Yaskawa INFORM job: 1.JBI

/JOB
//NAME 1
//POS
///NPOS 162,162,162,0,0,0
///TOOL 0
///POSTYPE PULSE
///PULSE
C00000=-283,-101162,-84213,3710,-80188,-1936
C00001=-283,-101162,-84213,3710,-80188,-1936
C00002=115939,-17843,-44700,-6904,-63515,59085
C00003=117709,3731,-51645,-6384,-54030,83191
C00004=117709,3731,-51645,-6384,-54030,83191
C00005=124817,11091,-45240,2225,-58232,65802
C00006=128558,-4341,-61499,8943,-39416,48451
C00007=141937,23059,-44881,39121,-57053,20454
C00008=142920,35333,-35255,42486,-63609,8178
C00009=131389,51659,-10555,16038,-74664,11710
C00010=126196,50041,-9511,12612,-72523,-6101
C00011=114039,49083,-11086,-6822,-73270,-17046
C00012=112111,54426,-8133,-7185,-80829,-32375
C00013=101553,48559,-20697,-28143,-77568,-33966
C00014=105123,31884,-31701,-21046,-69946,-46894
C00015=111650,18447,-39836,-11003,-63489,-61522
C00016=113485,7970,-48571,-14105,-57851,-74639
C00017=113485,7970,-48571,-14105,-57851,-74639
C00018=114170,-2374,-36949,-11645,-74681,-76938
C00019=113314,-7643,-38017,-11019,-76954,88145
C00020=102960,15783,-40712,-5055,-61801,87407
C00021=102960,15783,-40712,-5055,-61801,87407
C00022=109484,11848,-44448,3017,-57913,70801
C00023=111825,-4491,-61766,4155,-38221,55572
C00024=127233,18004,-49993,42137,-51406,23800
C00025=123794,20070,-44223,34245,-49783,15146
C00026=118261,52920,-9530,17828,-74428,15725
C00027=113721,45593,-13485,15354,-67043,-2855
C00028=99817,50806,-8879,-9234,-71758,-11440
C00029=100311,60695,-910,-3132,-82683,-29064
C00030=89808,58501,-9489,-23508,-82083,-31436
C00031=93781,55410,-9430,-14151,-84882,-46382
C00032=94766,20128,-39423,-16116,-61452,-54210
C00033=98573,11657,-45494,-13692,-58332,-69623
C00034=98573,11657,-45494,-13692,-58332,-69623
C00035=99303,8604,-31154,-10952,-72489,-71699
C00036=89422,16015,-23794,-2157,-75183,91094
C00037=90041,28841,-28187,-2386,-65884,91066
C00038=90041,28841,-28187,-2386,-65884,91066
C00039=95426,19332,-37606,3682,-57792,75417
C00040=103247,16005,-44070,17550,-50613,56089
C00041=113549,16841,-53361,50996,-44891,24333
C00042=112114,26764,-40359,41262,-49930,18196
C00043=105423,50717,-10337,19910,-67719,16523
C00044=102098,58112,-1142,17447,-71662,1302
C00045=90776,64198,5929,-1117,-76945,-10230
C00046=87727,74947,14485,-3611,-87418,-24219
C00047=79354,72723,7405,-19240,-87200,-29236
C00048=76420,55305,-10510,-24564,-76474,-35505
C00049=83670,16895,-41951,-12582,-49930,-51607
C00050=85054,23740,-34298,-12468,-60756,-65460
C00051=85054,23740,-34298,-12468,-60756,-65460
C00052=85063,22114,-18753,-9149,-74798,-67250
C00053=72786,31521,-9549,-9445,-75352,93043
C00054=77617,39381,-17527,-2945,-63917,95499
C00055=77617,39381,-17527,-2945,-63917,95499
C00056=81845,27264,-30649,1079,-52677,78149
C00057=86990,13258,-48946,12655,-33027,60150
C00058=90994,9633,-56784,33436,-24362,42962
C00059=99247,25142,-45272,51284,-40942,28841
C00060=98491,33379,-33635,41928,-45438,21477
C00061=97892,43719,-21091,40448,-51711,6672
C00062=90154,66189,8945,17735,-69591,4970
C00063=76670,80759,24898,-8994,-81212,-4057
C00064=77890,93073,36819,-863,-92684,-21133
C00065=70280,91760,31185,-15532,-93504,-27367
C00066=65704,69069,5703,-24854,-77527,-31557
C00067=69263,47501,-12611,-17938,-65429,-45438
C00068=73833,39987,-17909,-11044,-63928,-62173
C00069=73833,39987,-17909,-11044,-63928,-62173
C00070=75039,37514,-3449,-7701,-77257,-64173
C00071=74616,28156,-12897,-9694,-74827,92488
C00072=73614,40170,-17462,-11390,-64426,94165
C00073=73614,40170,-17462,-11390,-64426,94165
C00074=73614,40170,-17462,-11390,-64426,94165
C00075=81727,26723,-31141,1076,-52650,80628
C00076=86883,12521,-49454,12588,-33076,60218
C00077=90994,9713,-56809,33527,-24311,42932
C00078=90994,9713,-56809,33527,-24311,42932
C00079=99183,24902,-45504,51304,-40911,28852
C00080=99183,24902,-45504,51304,-40911,28852
C00081=98411,33440,-33412,41862,-45487,21541
C00082=99416,42526,-24620,46864,-51095,3725
C00083=90863,70401,13127,18633,-73267,4997
C00084=76675,81176,25590,-8988,-81419,-4073
C00085=77890,93045,36838,-863,-92708,-21133
C00086=70280,91719,31202,-15533,-93535,-27371
C00087=65715,68855,5477,-24835,-77499,-31559
C00088=66119,47846,-14846,-25675,-64947,-43795
C00089=70910,45228,-13849,-14534,-65052,-50806
C00090=75926,27198,-30687,-6609,-51803,-64018
C00091=75926,27198,-30687,-6609,-51803,-64018
C00092=74844,35432,-1015,-7610,-79822,-64270
C00093=74616,28156,-12897,-9694,-74827,92488
C00094=90411,-2677,-20047,-11125,-84138,86440
C00095=90413,-2674,-20051,-11105,-84138,86441
C00096=137757,-12075,-30464,2646,-72394,74401
C00097=139263,-65150,-85436,14259,-28990,73053
C00098=137079,-26031,-69593,36686,-11816,62677
C00099=137079,-26031,-69593,36686,-11816,62677
C00100=139435,-23870,-66142,38084,-15914,40453
C00101=138383,-26116,-69231,45202,-10210,18865
C00102=136988,-21816,-61713,19512,-16285,9124
C00103=134481,-8714,-45390,4049,-32022,-3278
C00104=132816,-12054,-49266,2863,-29473,-26222
C00105=133118,-16915,-54850,5104,-25691,-47193
C00106=132429,-23928,-65383,-2979,-14980,-66671
C00107=133899,-27903,-74314,23479,-2636,-94546
C00108=138833,-79965,-103111,19688,-12213,-93629
C00109=119564,-93872,-103655,-3232,-19191,84847
C00110=119617,-28274,-68464,-3848,-15128,84753
C00111=119617,-28274,-68464,-3848,-15128,84753
C00112=119575,-30245,-73045,-30117,-7907,72568
C00113=119533,-30199,-72935,-30139,-8105,72141
C00114=119084,-28019,-67713,-21117,-14338,49832
C00115=119103,-25674,-64433,-15990,-16239,28421
C00116=117904,-24651,-63335,-18016,-16610,10465
C00117=116364,-17323,-54707,-12430,-26691,-16379
C00118=116034,-19270,-56740,-12888,-26506,-35915
C00119=108922,-18911,-60992,-47912,-30029,-42936
C00120=114993,-30399,-76205,-74620,-10810,-47413
C00121=113126,-78683,-102705,-45607,-16425,-60367
C00122=119564,-93872,-103655,-3232,-19191,84847
C00123=119501,-30079,-72867,-7033,-8758,86614
C00124=119501,-30079,-72867,-7033,-8758,86614
C00125=119390,-30716,-74067,-37591,-7172,75727
C00126=121229,-29061,-69555,-4595,-11344,43979
C00127=119104,-25703,-64453,-15989,-16243,28419
C00128=118126,-13614,-49952,-9217,-30446,5536
C00129=116206,-13809,-50361,-10582,-31136,-17197
C00130=117334,-18567,-55575,-6506,-27346,-35991
C00131=112042,-24638,-66931,-46893,-21308,-43852
C00132=114210,-29455,-74183,-63406,-12970,-50800
C00133=113074,-79856,-103225,-44998,-16651,-60643
C00134=119564,-93872,-105617,-3232,-19191,84847
C00135=119749,-29508,-71257,-4806,-11297,85540
C00136=119749,-29508,-71257,-4806,-11297,85540
C00137=117863,-29016,-70107,-32919,-13598,71537
C00138=121387,-23775,-62079,-1920,-20330,42797
C00139=119104,-25781,-64508,-15983,-16250,28419
C00140=117899,-24917,-63521,-18002,-16633,10461
C00141=116021,-17584,-54917,-12768,-26744,-16159
C00142=113094,-17565,-56131,-24726,-28094,-26210
C00143=114237,-26152,-67609,-36989,-17763,-46723
C00144=115048,-30330,-76182,-74696,-10772,-47388
C00145=112648,-89264,-107216,-40476,-18619,-62704
C00146=119564,-93872,-105617,-3232,-19191,84847
C00147=119728,-31105,-75415,-11420,-5001,88504
C00148=119728,-31105,-75415,-11420,-5001,88504
C00149=120343,-30953,-74249,-21828,-6042,69534
C00150=126312,-14750,-51708,17407,-33389,37991
C00151=119102,-25993,-64654,-15969,-16267,28412
C00152=117899,-25020,-63592,-17997,-16641,10457
C00153=116085,-17534,-54630,-12641,-26883,-16232
C00154=116220,-19444,-56979,-12194,-26346,-35772
C00155=115970,-21766,-59500,-15760,-26236,-55559
C00156=114981,-30317,-76177,-74755,-10811,-47349
C00157=112538,-91654,-108181,-39431,-19159,-63177
C00158=112538,-91654,-78834,-11871,-48570,95336
C00159=112538,-91654,-78834,-11871,-48570,95336
C00160=-2476,-84373,-75976,-13540,-83606,15477
C00161=-283,-101162,-84213,3710,-80188,-1936
BC00000=570125
BC00001=868704
BC00002=878894
BC00003=878037
BC00004=878037
BC00005=878038
BC00006=878037
BC00007=878038
BC00008=878038
BC00009=878038
BC00010=878038
BC00011=878037
BC00012=878037
BC00013=878037
BC00014=878037
BC00015=878037
BC00016=878037
BC00017=878037
BC00018=878037
BC00019=912823
BC00020=878035
BC00021=878035
BC00022=878037
BC00023=878037
BC00024=878038
BC00025=878037
BC00026=878038
BC00027=878038
BC00028=878037
BC00029=878037
BC00030=878037
BC00031=878037
BC00032=878037
BC00033=878037
BC00034=878037
BC00035=878037
BC00036=878035
BC00037=878036
BC00038=878036
BC00039=878037
BC00040=878037
BC00041=878038
BC00042=878038
BC00043=878038
BC00044=878038
BC00045=878037
BC00046=878037
BC00047=878037
BC00048=878037
BC00049=878037
BC00050=878037
BC00051=878037
BC00052=878037
BC00053=878037
BC00054=878035
BC00055=878035
BC00056=877203
BC00057=877947
BC00058=878201
BC00059=878342
BC00060=878784
BC00061=877961
BC00062=877604
BC00063=878505
BC00064=878840
BC00065=878535
BC00066=877953
BC00067=879795
BC00068=878428
BC00069=878428
BC00070=878037
BC00071=915550
BC00072=913919
BC00073=913919
BC00074=913919
BC00075=916409
BC00076=916569
BC00077=916479
BC00078=916479
BC00079=916387
BC00080=916387
BC00081=916586
BC00082=915550
BC00083=915870
BC00084=916359
BC00085=916889
BC00086=917058
BC00087=916344
BC00088=917145
BC00089=916666
BC00090=915811
BC00091=915811
BC00092=915811
BC00093=915550
BC00094=915550
BC00095=915550
BC00096=915550
BC00097=915550
BC00098=915550
BC00099=915550
BC00100=915550
BC00101=915550
BC00102=915550
BC00103=915550
BC00104=915550
BC00105=915550
BC00106=915550
BC00107=915550
BC00108=915550
BC00109=915550
BC00110=915550
BC00111=915550
BC00112=915550
BC00113=915550
BC00114=915550
BC00115=915550
BC00116=915550
BC00117=915550
BC00118=915550
BC00119=915550
BC00120=915550
BC00121=915550
BC00122=954211
BC00123=953187
BC00124=953187
BC00125=954162
BC00126=953948
BC00127=954071
BC00128=953633
BC00129=953244
BC00130=953645
BC00131=954029
BC00132=953749
BC00133=953683
BC00134=992214
BC00135=992214
BC00136=992214
BC00137=991968
BC00138=992423
BC00139=992186
BC00140=992082
BC00141=991168
BC00142=991569
BC00143=992735
BC00144=991845
BC00145=991844
BC00146=1026906
BC00147=1030289
BC00148=1030289
BC00149=1030261
BC00150=1030281
BC00151=1030485
BC00152=1029902
BC00153=1029299
BC00154=1030152
BC00155=1030177
BC00156=1030552
BC00157=1030552
BC00158=1030552
BC00159=1030552
BC00160=952617
BC00161=570125
EC00000=1166,0
EC00001=1166,0
EC00002=-1742,0
EC00003=-1741,0
EC00004=-1741,0
EC00005=-1743,0
EC00006=-1742,0
EC00007=-1741,0
EC00008=-1741,0
EC00009=-1741,0
EC00010=-1741,0
EC00011=-1741,0
EC00012=-1741,0
EC00013=-1742,0
EC00014=-1742,0
EC00015=-1742,0
EC00016=-1741,0
EC00017=-1741,0
EC00018=-1741,0
EC00019=-1741,0
EC00020=-1744,0
EC00021=-1744,0
EC00022=-1742,0
EC00023=-1742,0
EC00024=-1741,0
EC00025=-1741,0
EC00026=-1741,0
EC00027=-1741,0
EC00028=-1741,0
EC00029=-1741,0
EC00030=-1742,0
EC00031=-1742,0
EC00032=-1741,0
EC00033=-1741,0
EC00034=-1741,0
EC00035=-1741,0
EC00036=-1743,0
EC00037=-1742,0
EC00038=-1742,0
EC00039=-1742,0
EC00040=-1742,0
EC00041=-1741,0
EC00042=-1741,0
EC00043=-1595,0
EC00044=-1742,0
EC00045=-1741,0
EC00046=-1741,0
EC00047=-1742,0
EC00048=-1742,0
EC00049=-1741,0
EC00050=-1741,0
EC00051=-1741,0
EC00052=-1741,0
EC00053=-1741,0
EC00054=-1743,0
EC00055=-1743,0
EC00056=-1742,0
EC00057=-1743,0
EC00058=-1742,0
EC00059=-1741,0
EC00060=-1741,0
EC00061=-1742,0
EC00062=-1742,0
EC00063=-1742,0
EC00064=-1741,0
EC00065=-1741,0
EC00066=-1741,0
EC00067=-1741,0
EC00068=-1742,0
EC00069=-1742,0
EC00070=-1741,0
EC00071=-1741,0
EC00072=-1742,0
EC00073=-1742,0
EC00074=-1742,0
EC00075=-1742,0
EC00076=-1743,0
EC00077=-1742,0
EC00078=-1742,0
EC00079=-1741,0
EC00080=-1741,0
EC00081=-1740,0
EC00082=-1742,0
EC00083=-1742,0
EC00084=-1742,0
EC00085=-1741,0
EC00086=-1741,0
EC00087=-1741,0
EC00088=-1742,0
EC00089=-1742,0
EC00090=-1742,0
EC00091=-1742,0
EC00092=-1741,0
EC00093=-1741,0
EC00094=-1741,0
EC00095=-84878,0
EC00096=-84879,0
EC00097=-84877,0
EC00098=-84877,0
EC00099=-84877,0
EC00100=-84877,0
EC00101=-84877,0
EC00102=-84877,0
EC00103=-84877,0
EC00104=-84877,0
EC00105=-84877,0
EC00106=-84877,0
EC00107=-84877,0
EC00108=-84877,0
EC00109=-84877,0
EC00110=-84877,0
EC00111=-84877,0
EC00112=-84877,0
EC00113=-84877,0
EC00114=-84877,0
EC00115=-84877,0
EC00116=-84877,0
EC00117=-84877,0
EC00118=-84877,0
EC00119=-84877,0
EC00120=-84877,0
EC00121=-84877,0
EC00122=-84877,0
EC00123=-84877,0
EC00124=-84877,0
EC00125=-84877,0
EC00126=-84877,0
EC00127=-84877,0
EC00128=-84877,0
EC00129=-84877,0
EC00130=-84877,0
EC00131=-84877,0
EC00132=-84877,0
EC00133=-84877,0
EC00134=-84877,0
EC00135=-84877,0
EC00136=-84877,0
EC00137=-84877,0
EC00138=-84877,0
EC00139=-84877,0
EC00140=-84877,0
EC00141=-84877,0
EC00142=-84877,0
EC00143=-84877,0
EC00144=-84877,0
EC00145=-84877,0
EC00146=-84877,0
EC00147=-84877,0
EC00148=-84877,0
EC00149=-84877,0
EC00150=-84877,0
EC00151=-84877,0
EC00152=-84877,0
EC00153=-84877,0
EC00154=-84877,0
EC00155=-84877,0
EC00156=-84877,0
EC00157=-84877,0
EC00158=-84877,0
EC00159=-2299,0
EC00160=-193,0
EC00161=1166,0
//INST
///DATE 2024/12/23 09:51
///COMM OZZ
///ATTR SC,RW
///GROUP1 RB1,BS1
///GROUP2 ST1
NOP
MOVJ C00000 BC00000 VJ=70.00 DEC=20  +MOVJ EC00000 VJ=70.00
MOVJ C00001 BC00001 VJ=40.00 DEC=20  +MOVJ EC00001 VJ=40.00
MOVJ C00002 BC00002 VJ=70.00 DEC=20  +MOVJ EC00002 VJ=70.00
MOVJ C00003 BC00003 VJ=40.00 DEC=20  +MOVJ EC00003 VJ=70.00
MACRO1 MJ#(0) ARGF5
ARCON
MOVC C00004 BC00004 V=4.2 DEC=20  +MOVJ EC00004 VJ=70.00
MOVC C00005 BC00005 V=4.2 DEC=20  +MOVJ EC00005 VJ=30.00
MOVC C00006 BC00006 V=4.2 DEC=20  +MOVJ EC00006 VJ=30.00
MOVC C00007 BC00007 V=4.2 DEC=20  +MOVJ EC00007 VJ=30.00
MOVC C00008 BC00008 V=4.2 DEC=20  +MOVJ EC00008 VJ=30.00
MOVC C00009 BC00009 V=4.2 DEC=20  +MOVJ EC00009 VJ=30.00
MOVC C00010 BC00010 V=4.2 DEC=20  +MOVJ EC00010 VJ=30.00
MOVC C00011 BC00011 V=4.2 DEC=20  +MOVJ EC00011 VJ=30.00
MOVC C00012 BC00012 V=4.2 DEC=20  +MOVJ EC00012 VJ=30.00
MOVC C00013 BC00013 V=4.2 DEC=20  +MOVJ EC00013 VJ=30.00
MOVC C00014 BC00014 V=4.2 DEC=20  +MOVJ EC00014 VJ=30.00
MOVC C00015 BC00015 V=4.2 DEC=20  +MOVJ EC00015 VJ=30.00
MOVC C00016 BC00016 V=4.2 DEC=20  +MOVJ EC00016 VJ=30.00
MOVJ C00017 BC00017 VJ=30.00 DEC=20  +MOVJ EC00017 VJ=30.00
ARCOF
MOVJ C00018 BC00018 VJ=40.00 DEC=20  +MOVJ EC00018 VJ=40.00
MOVJ C00019 BC00019 VJ=70.00 DEC=20  +MOVJ EC00019 VJ=0.78
MOVJ C00020 BC00020 VJ=30.00 DEC=20  +MOVJ EC00020 VJ=0.78
ARCON
MOVC C00021 BC00021 V=4.2 DEC=20  +MOVJ EC00021 VJ=0.78
MOVC C00022 BC00022 V=4.2 DEC=20  +MOVJ EC00022 VJ=0.78
MOVC C00023 BC00023 V=4.2 DEC=20  +MOVJ EC00023 VJ=30.00
MOVC C00024 BC00024 V=4.2 DEC=20  +MOVJ EC00024 VJ=30.00
MOVC C00025 BC00025 V=5.8 DEC=20  +MOVJ EC00025 VJ=30.00
MOVC C00026 BC00026 V=4.2 DEC=20  +MOVJ EC00026 VJ=30.00
MOVC C00027 BC00027 V=4.2 DEC=20  +MOVJ EC00027 VJ=30.00
MOVC C00028 BC00028 V=4.2 DEC=20  +MOVJ EC00028 VJ=30.00
MOVC C00029 BC00029 V=4.2 DEC=20  +MOVJ EC00029 VJ=30.00
MOVC C00030 BC00030 V=4.2 DEC=20  +MOVJ EC00030 VJ=30.00
MOVC C00031 BC00031 V=4.2 DEC=20  +MOVJ EC00031 VJ=30.00
MOVC C00032 BC00032 V=4.2 DEC=20  +MOVJ EC00032 VJ=30.00
MOVC C00033 BC00033 V=4.2 DEC=20  +MOVJ EC00033 VJ=30.00
MOVJ C00034 BC00034 VJ=25.00 DEC=20  +MOVJ EC00034 VJ=30.00
ARCOF
MOVJ C00035 BC00035 VJ=30.00 DEC=20  +MOVJ EC00035 VJ=30.00
MOVJ C00036 BC00036 VJ=30.00 DEC=20  +MOVJ EC00036 VJ=30.00
MOVJ C00037 BC00037 VJ=30.00 DEC=20  +MOVJ EC00037 VJ=30.00
ARCON
MOVC C00038 BC00038 V=4.2 DEC=20  +MOVJ EC00038 VJ=30.00
MOVC C00039 BC00039 V=4.2 DEC=20  +MOVJ EC00039 VJ=30.00
MOVC C00040 BC00040 V=4.2 DEC=20  +MOVJ EC00040 VJ=30.00
MOVC C00041 BC00041 V=4.2 DEC=20  +MOVJ EC00041 VJ=30.00
MOVC C00042 BC00042 V=4.2 DEC=20  +MOVJ EC00042 VJ=30.00
MOVC C00043 BC00043 V=4.2 DEC=20  +MOVJ EC00043 VJ=30.00
MOVC C00044 BC00044 V=4.2 DEC=20  +MOVJ EC00044 VJ=30.00
MOVC C00045 BC00045 V=4.2 DEC=20  +MOVJ EC00045 VJ=30.00
MOVC C00046 BC00046 V=4.2 DEC=20  +MOVJ EC00046 VJ=30.00
MOVC C00047 BC00047 V=4.2 DEC=20  +MOVJ EC00047 VJ=30.00
MOVC C00048 BC00048 V=5.8 DEC=20  +MOVJ EC00048 VJ=30.00
MOVC C00049 BC00049 V=4.2 DEC=20  +MOVJ EC00049 VJ=0.78
MOVC C00050 BC00050 V=4.2 DEC=20  +MOVJ EC00050 VJ=30.00
MOVJ C00051 BC00051 VJ=30.00 DEC=20  +MOVJ EC00051 VJ=30.00
ARCOF
MOVJ C00052 BC00052 VJ=30.00 DEC=20  +MOVJ EC00052 VJ=30.00
MOVJ C00053 BC00053 VJ=30.00 DEC=20  +MOVJ EC00053 VJ=30.00
MOVJ C00054 BC00054 VJ=30.00 DEC=20  +MOVJ EC00054 VJ=30.00
ARCON
MOVC C00055 BC00055 V=4.2 DEC=20  +MOVJ EC00055 VJ=30.00
MOVC C00056 BC00056 V=4.2 DEC=20  +MOVJ EC00056 VJ=0.78
MOVC C00057 BC00057 V=4.2 DEC=20  +MOVJ EC00057 VJ=0.78
MOVC C00058 BC00058 V=4.2 DEC=20  +MOVJ EC00058 VJ=0.78
MOVC C00059 BC00059 V=4.2 DEC=20  +MOVJ EC00059 VJ=0.78
MOVC C00060 BC00060 V=4.2 DEC=20  +MOVJ EC00060 VJ=0.78
MOVC C00061 BC00061 V=4.2 DEC=20  +MOVJ EC00061 VJ=0.78
MOVC C00062 BC00062 V=4.2 DEC=20  +MOVJ EC00062 VJ=0.78
MOVC C00063 BC00063 V=4.2 DEC=20  +MOVJ EC00063 VJ=0.78
MOVC C00064 BC00064 V=4.2 DEC=20  +MOVJ EC00064 VJ=0.78
MOVC C00065 BC00065 V=4.2 DEC=20  +MOVJ EC00065 VJ=0.78
MOVC C00066 BC00066 V=4.2 DEC=20  +MOVJ EC00066 VJ=0.78
MOVC C00067 BC00067 V=4.2 DEC=20  +MOVJ EC00067 VJ=0.78
MOVC C00068 BC00068 V=4.2 DEC=20  +MOVJ EC00068 VJ=0.78
MOVJ C00069 BC00069 VJ=30.00 DEC=20  +MOVJ EC00069 VJ=30.00
ARCOF
MOVJ C00070 BC00070 VJ=30.00 DEC=20  +MOVJ EC00070 VJ=30.00
MOVJ C00071 BC00071 VJ=30.00 DEC=20  +MOVJ EC00071 VJ=30.00
MOVJ C00072 BC00072 VJ=30.00 DEC=20  +MOVJ EC00072 VJ=30.00
MOVC C00073 BC00073 V=116.7 DEC=20  +MOVJ EC00073 VJ=0.78
ARCON
MOVC C00074 BC00074 V=4.2 DEC=20  +MOVJ EC00074 VJ=30.00
MOVC C00075 BC00075 V=4.2 DEC=20  +MOVJ EC00075 VJ=30.00
MOVC C00076 BC00076 V=4.2 DEC=20  +MOVJ EC00076 VJ=30.00
MOVC C00077 BC00077 V=4.2 DEC=20  +MOVJ EC00077 VJ=40.00
MOVJ C00078 BC00078 VJ=70.00 DEC=20  +MOVJ EC00078 VJ=70.00
MOVC C00079 BC00079 V=4.2 DEC=20  +MOVJ EC00079 VJ=30.00
MOVC C00080 BC00080 V=4.2 DEC=20  +MOVJ EC00080 VJ=25.00
MOVC C00081 BC00081 V=4.2 DEC=20  +MOVJ EC00081 VJ=25.00
MOVC C00082 BC00082 V=4.2 DEC=20  +MOVJ EC00082 VJ=30.00
MOVC C00083 BC00083 V=4.2 DEC=20  +MOVJ EC00083 VJ=70.00
MOVC C00084 BC00084 V=4.2 DEC=20  +MOVJ EC00084 VJ=30.00
MOVC C00085 BC00085 V=4.2 DEC=20  +MOVJ EC00085 VJ=30.00
MOVC C00086 BC00086 V=4.2 DEC=20  +MOVJ EC00086 VJ=30.00
MOVC C00087 BC00087 V=4.2 DEC=20  +MOVJ EC00087 VJ=30.00
MOVC C00088 BC00088 V=4.2 DEC=20  +MOVJ EC00088 VJ=30.00
MOVC C00089 BC00089 V=4.2 DEC=20  +MOVJ EC00089 VJ=0.78
MOVC C00090 BC00090 V=4.2 DEC=20  +MOVJ EC00090 VJ=30.00
MOVJ C00091 BC00091 VJ=25.00 DEC=20  +MOVJ EC00091 VJ=30.00
ARCOF
MOVJ C00092 BC00092 VJ=30.00 DEC=20  +MOVJ EC00092 VJ=30.00
MOVJ C00093 BC00093 VJ=30.00 DEC=20  +MOVJ EC00093 VJ=30.00
MOVJ C00094 BC00094 VJ=30.00 DEC=20  +MOVJ EC00094 VJ=30.00
MOVJ C00095 BC00095 VJ=30.00 DEC=20  +MOVJ EC00095 VJ=30.00
MOVJ C00096 BC00096 VJ=30.00 DEC=20  +MOVJ EC00096 VJ=30.00
MOVJ C00097 BC00097 VJ=0.78 DEC=20  +MOVJ EC00097 VJ=0.78
MOVJ C00098 BC00098 VJ=30.00 DEC=20  +MOVJ EC00098 VJ=0.78
ARCON
MOVC C00099 BC00099 V=5.0 DEC=20  +MOVJ EC00099 VJ=0.78
MOVC C00100 BC00100 V=5.0 DEC=20  +MOVJ EC00100 VJ=0.78
MOVC C00101 BC00101 V=5.0 DEC=20  +MOVJ EC00101 VJ=0.78
MOVC C00102 BC00102 V=5.0 DEC=20  +MOVJ EC00102 VJ=0.78
MOVC C00103 BC00103 V=5.0 DEC=20  +MOVJ EC00103 VJ=0.78
MOVC C00104 BC00104 V=5.0 DEC=20  +MOVJ EC00104 VJ=0.78
MOVC C00105 BC00105 V=5.0 DEC=20  +MOVJ EC00105 VJ=0.78
MOVC C00106 BC00106 V=5.0 DEC=20  +MOVJ EC00106 VJ=0.78
MOVC C00107 BC00107 V=5.0 DEC=20  +MOVJ EC00107 VJ=0.78
ARCOF
MOVJ C00108 BC00108 VJ=40.00 DEC=20  +MOVJ EC00108 VJ=0.78
MOVJ C00109 BC00109 VJ=40.00 DEC=20  +MOVJ EC00109 VJ=0.78
MOVJ C00110 BC00110 VJ=40.00 DEC=20  +MOVJ EC00110 VJ=0.78
ARCON
MOVC C00111 BC00111 V=5.0 DEC=20  +MOVJ EC00111 VJ=0.78
MOVC C00112 BC00112 V=5.0 DEC=20  +MOVJ EC00112 VJ=0.78
MOVC C00113 BC00113 V=5.0 DEC=20  +MOVJ EC00113 VJ=0.78
MOVC C00114 BC00114 V=5.0 DEC=20  +MOVJ EC00114 VJ=40.00
MOVC C00115 BC00115 V=5.0 DEC=20  +MOVJ EC00115 VJ=0.78
MOVC C00116 BC00116 V=5.0 DEC=20  +MOVJ EC00116 VJ=0.78
MOVC C00117 BC00117 V=5.0 DEC=20  +MOVJ EC00117 VJ=0.78
MOVC C00118 BC00118 V=5.0 DEC=20  +MOVJ EC00118 VJ=0.78
MOVC C00119 BC00119 V=5.0 DEC=20  +MOVJ EC00119 VJ=0.78
MOVC C00120 BC00120 V=5.0 DEC=20  +MOVJ EC00120 VJ=0.78
ARCOF
MOVJ C00121 BC00121 VJ=40.00 DEC=20  +MOVJ EC00121 VJ=0.78
MOVJ C00122 BC00122 VJ=40.00 DEC=20  +MOVJ EC00122 VJ=0.78
MOVJ C00123 BC00123 VJ=40.00 DEC=20  +MOVJ EC00123 VJ=0.78
ARCON
MOVC C00124 BC00124 V=5.0 DEC=20  +MOVJ EC00124 VJ=0.78
MOVC C00125 BC00125 V=5.0 DEC=20  +MOVJ EC00125 VJ=0.78
MOVC C00126 BC00126 V=5.0 DEC=20  +MOVJ EC00126 VJ=0.78
MOVC C00127 BC00127 V=5.0 DEC=20  +MOVJ EC00127 VJ=0.78
MOVC C00128 BC00128 V=5.0 DEC=20  +MOVJ EC00128 VJ=0.78
MOVC C00129 BC00129 V=5.0 DEC=20  +MOVJ EC00129 VJ=0.78
MOVC C00130 BC00130 V=5.0 DEC=20  +MOVJ EC00130 VJ=0.78
MOVC C00131 BC00131 V=5.0 DEC=20  +MOVJ EC00131 VJ=0.78
MOVC C00132 BC00132 V=5.0 DEC=20  +MOVJ EC00132 VJ=0.78
ARCOF
MOVJ C00133 BC00133 VJ=40.00 DEC=20  +MOVJ EC00133 VJ=0.78
MOVJ C00134 BC00134 VJ=40.00 DEC=20  +MOVJ EC00134 VJ=0.78
MOVJ C00135 BC00135 VJ=40.00 DEC=20  +MOVJ EC00135 VJ=0.78
ARCON
MOVC C00136 BC00136 V=5.0 DEC=20  +MOVJ EC00136 VJ=0.78
MOVC C00137 BC00137 V=5.0 DEC=20  +MOVJ EC00137 VJ=0.78
MOVC C00138 BC00138 V=5.0 DEC=20  +MOVJ EC00138 VJ=0.78
MOVC C00139 BC00139 V=5.0 DEC=20  +MOVJ EC00139 VJ=0.78
MOVC C00140 BC00140 V=5.0 DEC=20  +MOVJ EC00140 VJ=0.78
MOVC C00141 BC00141 V=5.0 DEC=20  +MOVJ EC00141 VJ=0.78
MOVC C00142 BC00142 V=5.0 DEC=20  +MOVJ EC00142 VJ=0.78
MOVC C00143 BC00143 V=5.0 DEC=20  +MOVJ EC00143 VJ=0.78
MOVC C00144 BC00144 V=5.0 DEC=20  +MOVJ EC00144 VJ=0.78
ARCOF
MOVJ C00145 BC00145 VJ=40.00 DEC=20  +MOVJ EC00145 VJ=0.78
MOVJ C00146 BC00146 VJ=40.00 DEC=20  +MOVJ EC00146 VJ=0.78
MOVJ C00147 BC00147 VJ=40.00 DEC=20  +MOVJ EC00147 VJ=0.78
ARCON
MOVC C00148 BC00148 V=5.0 DEC=20  +MOVJ EC00148 VJ=0.78
MOVC C00149 BC00149 V=5.0 DEC=20  +MOVJ EC00149 VJ=0.78
MOVC C00150 BC00150 V=5.0 DEC=20  +MOVJ EC00150 VJ=0.78
MOVC C00151 BC00151 V=5.0 DEC=20  +MOVJ EC00151 VJ=0.78
MOVC C00152 BC00152 V=5.0 DEC=20  +MOVJ EC00152 VJ=0.78
MOVC C00153 BC00153 V=5.0 DEC=20  +MOVJ EC00153 VJ=0.78
MOVC C00154 BC00154 V=5.0 DEC=20  +MOVJ EC00154 VJ=0.78
MOVC C00155 BC00155 V=5.0 DEC=20  +MOVJ EC00155 VJ=0.78
MOVC C00156 BC00156 V=5.0 DEC=20  +MOVJ EC00156 VJ=0.78
ARCOF
MOVJ C00157 BC00157 VJ=40.00 DEC=20  +MOVJ EC00157 VJ=0.78
MOVJ C00158 BC00158 VJ=40.00 DEC=20  +MOVJ EC00158 VJ=0.78
MOVJ C00159 BC00159 VJ=40.00 DEC=20  +MOVJ EC00159 VJ=40.00
MOVJ C00160 BC00160 VJ=40.00 DEC=20  +MOVJ EC00160 VJ=0.78
MOVJ C00161 BC00161 VJ=40.00 DEC=20  +MOVJ EC00161 VJ=0.78
END
